(* IEC 61131-3 sources: Gen-AI/final/Gen-AI_v1.0_submission/A2_框架源码/agent/logs/full34_fixture/E3_P06_1_42/tools/candidate_1/fixture_compile, 1 file *)

(* ---- source.st ---- *)
FUNCTION_BLOCK FB_P06
VAR_INPUT
    DO_LOW : BOOL;
    AERATION_E_STOP_NC : BOOL;
END_VAR
VAR_OUTPUT
    BLOWER_RUN : BOOL;
    AERATION_BLOWER_CYCLE_COUNT : UINT;
END_VAR
(* Add a VAR block for internal state/timers before the implementation, if needed. *)
(* SKELETON ONLY: replace this RETURN with scan logic and required initial state. *)
RETURN;
END_FUNCTION_BLOCK

(* FIXTURE_COMPILE_FAIL *)
